Staubli VAL3: _bindTRAJ.pgx

program _bindTRAJ()
  local num l_i
  local string l_sbtn
begin
  for l_i = 1 to 6
    l_sbtn="btn"+toString("",l_i)
    userPageBindClick("insertTRAJ",l_sbtn,bInsert[l_i],true)
  endFor

  userPageBind("insertTRAJ","lbl1","innerHTML",sPgIndexTRAJ,1,"r")
  userPageBind("insertTRAJ","lbl2","innerHTML",sPageTRAJ,1,"r")


  userPageBind("insertTRAJ","lst1","value",sInsertItem,1,"rw")
end
